Fanuc KAREL source: kt00108.KL

-- PROVISIONAL review KL for V1013-1; original PC SHA256 dbd1f374cac46ae093565d834c702cecc50c2da450888b1e9463e3d14fd033fe
-- Incomplete behavior may be omitted. Consult companion uncertainty JSON. Do not deploy.
PROGRAM KT00108
%NOLOCKGROUP
VAR
  R1 : REAL
  R2 : REAL
  OUT : REAL
BEGIN
  -- UNRESOLVED_PC offsets 5-16; opcodes 2E,23
  -- UNRESOLVED_PC offsets 21-32; opcodes 2E,23
  -- UNRESOLVED_PC offsets 37-48; opcodes 2E,23
  -- UNRESOLVED_PC offsets 53-64; opcodes 2E,23
  -- UNRESOLVED_PC offsets 69-88; opcodes 21,21,6C,23
  -- UNRESOLVED_PC offsets 93-97; opcodes 7F
END KT00108
